TYPE ST_8Bit :
STRUCT
    b0: BIT;
    b1: BIT;
    b2: BIT;
    b3: BIT;
    b4: BIT;
    b5: BIT;
    b6: BIT;
    b7: BIT;
END_STRUCT
END_TYPE

(* stored: Version 1.1.0.1
   DUT ST_8Bit: Id {48280b74-dab2-07cb-0277-17e101816ef4} *)
